ABB RAPID module: Main.mod

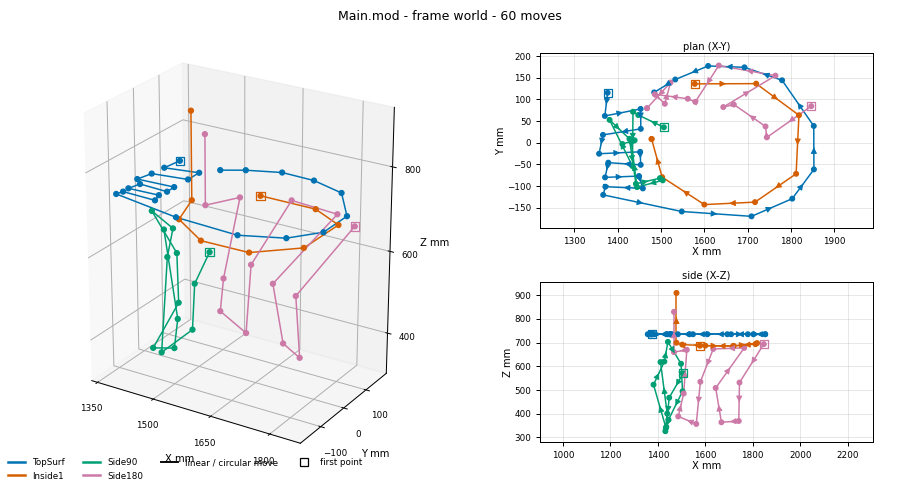
[picture p0: tool path of Main.mod in frame world, 60 of 82 moves have a stored position in this frame; points joined in program order, loops and branches not executed]
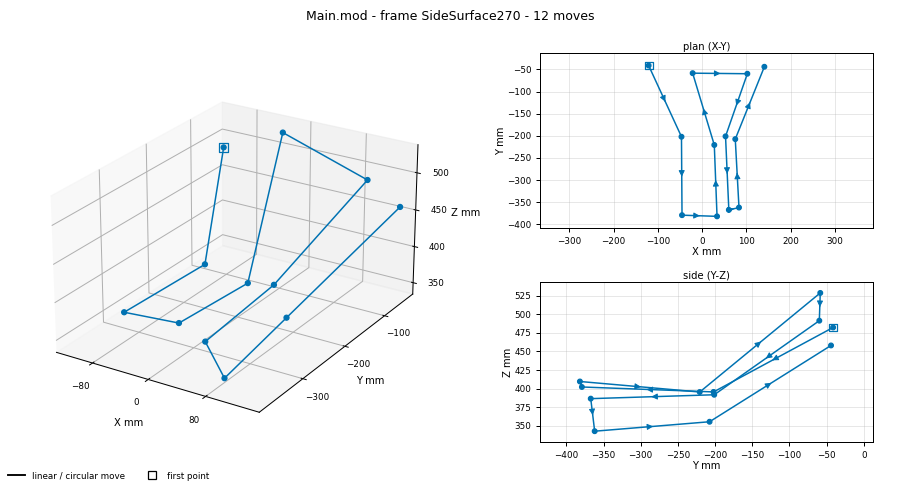
[picture p1: tool path of Main.mod in frame SideSurface270, 12 of 82 moves have a stored position in this frame; points joined in program order, loops and branches not executed]
%%%
  VERSION:1
  LANGUAGE:ENGLISH
%%%
MODULE MOD_Main

    ! -------------------------------
    ! Define customized variables here
    ! ...

	! Tool variables:
	PERS tooldata ToolRDK2 := [TRUE,[[-397.000,-4.578,191.692],[0.70710678,0.00000000,-0.70710678,0.00000001]],[1,[0,0,20],[1,0,0,0],0,0,0.005]];
	PERS tooldata ToolRDKRy15 := [TRUE,[[-327.000,-4.578,191.692],[0.60876143,0.00000000,-0.79335334,-0.00000000]],[1,[0,0,20],[1,0,0,0],0,0,0.005]];

	! Reference variables:
	PERS wobjdata SideSurface270 := [FALSE, TRUE, "", [[0,0,0],[1,0,0,0]],[[1336.130,0.000,735.410],[0.50000000,0.50000000,0.50000000,0.50000000]]];
	PERS wobjdata TopSurf2 := [FALSE, TRUE, "", [[0,0,0],[1,0,0,0]],[[1336.130,0.000,735.410],[0.50000000,0.50000000,0.50000000,0.50000000]]];
	PERS wobjdata Inside := [FALSE, TRUE, "", [[0,0,0],[1,0,0,0]],[[1336.130,0.000,735.410],[0.50000000,0.50000000,0.50000000,0.50000000]]];
	PERS wobjdata SideSurface90 := [FALSE, TRUE, "", [[0,0,0],[1,0,0,0]],[[1336.130,0.000,735.410],[0.50000000,0.50000000,0.50000000,0.50000000]]];
	PERS wobjdata SdeSurface180 := [FALSE, TRUE, "", [[0,0,0],[1,0,0,0]],[[1336.130,0.000,735.410],[0.50000000,0.50000000,0.50000000,0.50000000]]];

	PROC TopSurf()
		ConfJ \On;
		ConfL \Off;
		TT0deg;
		ToolRDK2 := [TRUE,[[-397.000,-4.578,191.692],[0.70710678,0.00000000,-0.70710678,0.00000001]],[1,[0,0,20],[1,0,0,0],0,0,0.005]];
		MoveAbsJ [[-2.762230,35.281600,-32.244600,94.063100,36.825000,84.928900],[9E+09,9E+09,9E+09,9E+09,9E+09,9E+09]],v500,z1,ToolRDK2 \WObj:=TopSurf2;
		MoveAbsJ [[3.888270,37.649400,-27.622300,84.244200,-60.438300,101.547000],[9E+09,9E+09,9E+09,9E+09,9E+09,9E+09]],v500,z1,ToolRDK2 \WObj:=TopSurf2;
		GunOn 1;
		MoveL [[115.290,-0.000,40.893],[0.66951661,0.66951663,0.22748073,-0.22748077],[-1,1,1,2],[9E+09,9E+09,9E+09,9E+09,9E+09,9E+09]],v500,z1,ToolRDK2 \WObj:=TopSurf2;
		MoveL [[61.769,-0.000,34.498],[0.66824739,0.66824741,0.23118262,-0.23118267],[0,0,1,1],[9E+09,9E+09,9E+09,9E+09,9E+09,9E+09]],v500,z1,ToolRDK2 \WObj:=TopSurf2;
		MoveL [[77.918,0.000,116.954],[0.67411479,0.67411479,0.21346957,-0.21346957],[0,0,1,1],[9E+09,9E+09,9E+09,9E+09,9E+09,9E+09]],v500,z1,ToolRDK2 \WObj:=TopSurf2;
		MoveL [[32.029,0.000,117.425],[0.67416339,0.67416339,0.21331602,-0.21331602],[0,0,1,1],[9E+09,9E+09,9E+09,9E+09,9E+09,9E+09]],v500,z1,ToolRDK2 \WObj:=TopSurf2;
		MoveL [[18.094,-0.000,30.124],[0.66795555,0.66795555,0.23202454,-0.23202454],[0,0,1,1],[9E+09,9E+09,9E+09,9E+09,9E+09,9E+09]],v500,z1,ToolRDK2 \WObj:=TopSurf2;
		MoveL [[-25.377,-0.000,21.201],[0.66687834,0.66687834,0.23510269,-0.23510270],[0,0,1,1],[9E+09,9E+09,9E+09,9E+09,9E+09,9E+09]],v500,z1,ToolRDK2 \WObj:=TopSurf2;
		MoveL [[-20.929,0.000,115.878],[0.67369753,0.67369752,0.21478279,-0.21478278],[0,0,1,1],[9E+09,9E+09,9E+09,9E+09,9E+09,9E+09]],v500,z1,ToolRDK2 \WObj:=TopSurf2;
		MoveL [[-51.029,0.000,117.232],[0.67365028,0.67365028,0.21493093,-0.21493093],[0,0,1,1],[9E+09,9E+09,9E+09,9E+09,9E+09,9E+09]],v500,z1,ToolRDK2 \WObj:=TopSurf2;
		MoveL [[-45.916,-0.000,42.441],[0.66826232,0.66826233,0.23113949,-0.23113950],[0,0,1,1],[9E+09,9E+09,9E+09,9E+09,9E+09,9E+09]],v500,z1,ToolRDK2 \WObj:=TopSurf2;
		MoveL [[-79.907,-0.000,34.972],[0.66736193,0.66736194,0.23372644,-0.23372644],[0,0,1,1],[9E+09,9E+09,9E+09,9E+09,9E+09,9E+09]],v500,z1,ToolRDK2 \WObj:=TopSurf2;
		MoveL [[-76.800,0.000,113.142],[0.67321469,0.67321469,0.21629141,-0.21629141],[0,0,1,1],[9E+09,9E+09,9E+09,9E+09,9E+09,9E+09]],v500,z1,ToolRDK2 \WObj:=TopSurf2;
		MoveL [[-105.332,0.000,122.191],[0.67370783,0.67370783,0.21475045,-0.21475045],[0,0,1,1],[9E+09,9E+09,9E+09,9E+09,9E+09,9E+09]],v500,z1,ToolRDK2 \WObj:=TopSurf2;
		MoveL [[-101.402,-0.000,35.713],[0.66719553,0.66719554,0.23420101,-0.23420104],[0,0,1,1],[9E+09,9E+09,9E+09,9E+09,9E+09,9E+09]],v500,z1,ToolRDK2 \WObj:=TopSurf2;
		MoveL [[-120.231,-0.000,30.646],[0.66659020,0.66659020,0.23591842,-0.23591844],[0,0,1,1],[9E+09,9E+09,9E+09,9E+09,9E+09,9E+09]],v500,z1,ToolRDK2 \WObj:=TopSurf2;
		MoveL [[-158.578,-0.000,211.837],[0.67989399,0.67989399,0.19427858,-0.19427858],[0,2,-1,0],[9E+09,9E+09,9E+09,9E+09,9E+09,9E+09]],v500,z1,ToolRDK2 \WObj:=TopSurf2;
		MoveL [[-169.769,-0.000,372.687],[0.68989069,0.68989069,0.15508330,-0.15508330],[0,2,-1,0],[9E+09,9E+09,9E+09,9E+09,9E+09,9E+09]],v500,z1,ToolRDK2 \WObj:=TopSurf2;
		MoveL [[-128.964,0.000,466.626],[0.69493868,0.69493868,0.13061485,-0.13061485],[0,2,-1,0],[9E+09,9E+09,9E+09,9E+09,9E+09,9E+09]],v500,z1,ToolRDK2 \WObj:=TopSurf2;
		MoveL [[-61.529,0.000,516.598],[0.69594843,0.69594843,0.12512308,-0.12512308],[0,2,-1,0],[9E+09,9E+09,9E+09,9E+09,9E+09,9E+09]],v500,z1,ToolRDK2 \WObj:=TopSurf2;
		MoveL [[38.647,0.000,516.273],[0.69521781,0.69521781,0.12912086,-0.12912086],[0,2,-1,0],[9E+09,9E+09,9E+09,9E+09,9E+09,9E+09]],v500,z1,ToolRDK2 \WObj:=TopSurf2;
		MoveL [[144.073,0.000,443.157],[0.69160511,0.69160511,0.14724934,-0.14724934],[0,0,1,1],[9E+09,9E+09,9E+09,9E+09,9E+09,9E+09]],v500,z1,ToolRDK2 \WObj:=TopSurf2;
		MoveL [[173.888,-0.000,356.448],[0.68759917,0.68759917,0.16494659,-0.16494659],[0,0,1,1],[9E+09,9E+09,9E+09,9E+09,9E+09,9E+09]],v500,z1,ToolRDK2 \WObj:=TopSurf2;
		MoveL [[177.057,0.000,272.670],[0.68344550,0.68344550,0.18138976,-0.18138976],[0,0,1,1],[9E+09,9E+09,9E+09,9E+09,9E+09,9E+09]],v500,z1,ToolRDK2 \WObj:=TopSurf2;
		MoveL [[145.838,-0.000,196.841],[0.67931130,0.67931130,0.19630627,-0.19630627],[0,0,1,1],[9E+09,9E+09,9E+09,9E+09,9E+09,9E+09]],v500,z1,ToolRDK2 \WObj:=TopSurf2;
		GunOn 0;
		MoveL [[116.077,0.000,148.259],[0.67637750,0.67637750,0.20618797,-0.20618797],[0,0,1,1],[9E+09,9E+09,9E+09,9E+09,9E+09,9E+09]],v500,z1,ToolRDK2 \WObj:=TopSurf2;
	ENDPROC

	PROC TT0deg()
		ConfJ \On;
		ConfL \Off;
		MoveAbsJ [[0.000000,0.000000,0.000000,0.000000,0.000000,0.000000],[9E+09,9E+09,9E+09,9E+09,9E+09,9E+09]],v500,z1,ToolRDK2 \WObj:=TopSurf2;
	ENDPROC

	PROC Inside1()
		ConfJ \On;
		ConfL \Off;
		TT0deg;
		MoveAbsJ [[-5.345720,35.456100,-20.669400,-15.550700,88.287700,-47.645500],[9E+09,9E+09,9E+09,9E+09,9E+09,9E+09]],v500,z1,ToolRDKRy15 \WObj:=Inside;
		GunOn 1;
		MoveL [[135.749,-48.253,241.842],[0.26164486,-0.62731638,0.51686708,-0.52044649],[-1,-1,-2,0],[9E+09,9E+09,9E+09,9E+09,9E+09,9E+09]],v100,z1,ToolRDKRy15 \WObj:=Inside;
		MoveL [[136.293,-48.875,383.457],[0.53837192,-0.31876420,0.47937269,-0.61542415],[-1,-1,3,0],[9E+09,9E+09,9E+09,9E+09,9E+09,9E+09]],v100,z1,ToolRDKRy15 \WObj:=Inside;
		MoveL [[63.451,-37.348,482.087],[0.60930435,-0.14318770,0.26615634,-0.73308001],[0,-1,3,0],[9E+09,9E+09,9E+09,9E+09,9E+09,9E+09]],v100,z1,ToolRDKRy15 \WObj:=Inside;
		MoveL [[-71.616,-41.647,475.560],[0.73598605,0.22123419,-0.09604572,-0.63257820],[-1,0,0,0],[9E+09,9E+09,9E+09,9E+09,9E+09,9E+09]],v100,z1,ToolRDKRy15 \WObj:=Inside;
		MoveL [[-136.962,-50.085,380.769],[0.64868094,0.45794626,-0.34884692,-0.49779925],[-1,0,0,0],[9E+09,9E+09,9E+09,9E+09,9E+09,9E+09]],v100,z1,ToolRDKRy15 \WObj:=Inside;
		MoveL [[-142.620,-47.996,263.919],[0.46214789,0.64281008,-0.47460814,-0.38465783],[-1,0,1,0],[9E+09,9E+09,9E+09,9E+09,9E+09,9E+09]],v100,z1,ToolRDKRy15 \WObj:=Inside;
		MoveL [[-79.374,-43.840,166.588],[0.24696012,0.71987130,-0.64178535,-0.09437996],[-1,0,1,0],[9E+09,9E+09,9E+09,9E+09,9E+09,9E+09]],v100,z1,ToolRDKRy15 \WObj:=Inside;
		MoveL [[8.609,-35.875,142.282],[0.04464887,0.71177006,-0.69465400,0.09405146],[-1,0,2,0],[9E+09,9E+09,9E+09,9E+09,9E+09,9E+09]],v100,z1,ToolRDKRy15 \WObj:=Inside;
		GunOn 0;
		MoveL [[8.609,174.125,142.282],[0.04464720,0.71176897,-0.69465549,0.09404953],[0,3,4,0],[9E+09,9E+09,9E+09,9E+09,9E+09,9E+09]],v100,z1,ToolRDKRy15 \WObj:=Inside;
	ENDPROC

	PROC Side90()
		ConfJ \On;
		ConfL \Off;
		TT90deg;
		ToolRDK2 := [TRUE,[[-397.000,-4.578,191.692],[0.70710678,0.00000000,-0.70710678,0.00000001]],[1,[0,0,20],[1,0,0,0],0,0,0.005]];
		MoveAbsJ [[2.579840,12.805000,8.075260,-0.378023,73.507000,3.846430],[9E+09,9E+09,9E+09,9E+09,9E+09,9E+09]],v100,z1,ToolRDK2 \WObj:=SideSurface90;
		MoveL [[35.648,-164.659,170.589],[0.70282661,0.03396154,0.01983662,-0.71027310],[0,-1,0,0],[9E+09,9E+09,9E+09,9E+09,9E+09,9E+09]],v100,z1,ToolRDK2 \WObj:=SideSurface90;
		GunOn 1;
		MoveL [[63.939,-267.719,111.565],[0.70282661,0.03396154,0.01983662,-0.71027310],[0,-1,0,0],[9E+09,9E+09,9E+09,9E+09,9E+09,9E+09]],v100,z1,ToolRDK2 \WObj:=SideSurface90;
		MoveL [[71.496,-390.187,99.400],[0.70282661,0.03396154,0.01983662,-0.71027310],[0,-1,0,0],[9E+09,9E+09,9E+09,9E+09,9E+09,9E+09]],v100,z1,ToolRDK2 \WObj:=SideSurface90;
		MoveL [[-53.749,-395.227,98.058],[0.70282661,0.03396154,0.01983662,-0.71027310],[-1,-1,0,0],[9E+09,9E+09,9E+09,9E+09,9E+09,9E+09]],v100,z1,ToolRDK2 \WObj:=SideSurface90;
		MoveL [[52.643,-212.764,45.439],[0.70282661,0.03396154,0.01983662,-0.71027310],[0,-1,0,0],[9E+09,9E+09,9E+09,9E+09,9E+09,9E+09]],v100,z1,ToolRDK2 \WObj:=SideSurface90;
		MoveL [[8.984,-115.328,91.184],[0.70282661,0.03396154,0.01983662,-0.71027310],[0,-1,0,0],[9E+09,9E+09,9E+09,9E+09,9E+09,9E+09]],v100,z1,ToolRDK2 \WObj:=SideSurface90;
		MoveL [[-94.720,-32.255,106.179],[0.70282661,0.03396154,0.01983662,-0.71027310],[-1,-1,-1,0],[9E+09,9E+09,9E+09,9E+09,9E+09,9E+09]],v100,z1,ToolRDK2 \WObj:=SideSurface90;
		MoveL [[-81.740,-124.404,161.457],[0.70282661,0.03396154,0.01983662,-0.71027310],[-1,-1,-1,0],[9E+09,9E+09,9E+09,9E+09,9E+09,9E+09]],v100,z1,ToolRDK2 \WObj:=SideSurface90;
		MoveL [[-86.756,-240.544,167.927],[0.70282661,0.03396154,0.01983662,-0.71027310],[-1,-1,-1,0],[9E+09,9E+09,9E+09,9E+09,9E+09,9E+09]],v100,z1,ToolRDK2 \WObj:=SideSurface90;
		MoveL [[-102.328,-360.623,108.637],[0.70282661,0.03396154,0.01983662,-0.71027310],[-1,-1,-1,0],[9E+09,9E+09,9E+09,9E+09,9E+09,9E+09]],v100,z1,ToolRDK2 \WObj:=SideSurface90;
		MoveL [[1.978,-408.957,95.385],[0.70282661,0.03396154,0.01983662,-0.71027310],[0,-1,0,0],[9E+09,9E+09,9E+09,9E+09,9E+09,9E+09]],v100,z1,ToolRDK2 \WObj:=SideSurface90;
		MoveL [[5.518,-334.746,103.233],[0.70282661,0.03396154,0.01983662,-0.71027310],[0,-1,0,0],[9E+09,9E+09,9E+09,9E+09,9E+09,9E+09]],v100,z1,ToolRDK2 \WObj:=SideSurface90;
		MoveL [[-2.937,-117.398,74.861],[0.70282661,0.03396154,0.01983662,-0.71027310],[0,-1,0,0],[9E+09,9E+09,9E+09,9E+09,9E+09,9E+09]],v100,z1,ToolRDK2 \WObj:=SideSurface90;
		GunOn 0;
	ENDPROC

	PROC TT90deg()
		ConfJ \On;
		ConfL \Off;
		MoveAbsJ [[90.000000,0.000000,0.000000,0.000000,0.000000,0.000000],[9E+09,9E+09,9E+09,9E+09,9E+09,9E+09]],v100,z1,ToolRDK2 \WObj:=SideSurface90;
	ENDPROC

	PROC Side180()
		ConfJ \On;
		ConfL \Off;
		TT180deg;
		ToolRDK2 := [TRUE,[[-397.000,-4.578,191.692],[0.70710678,0.00000000,-0.70710678,0.00000001]],[1,[0,0,20],[1,0,0,0],0,0,0.005]];
		MoveAbsJ [[22.186600,36.517800,-32.653500,15.382700,96.981900,81.677400],[9E+09,9E+09,9E+09,9E+09,9E+09,9E+09]],v100,z1,ToolRDK2 \WObj:=SdeSurface180;
		MoveL [[84.401,-41.748,510.527],[0.27194744,0.74951284,-0.59519100,-0.10011380],[-1,-1,-1,0],[9E+09,9E+09,9E+09,9E+09,9E+09,9E+09]],v100,z1,ToolRDK2 \WObj:=SdeSurface180;
		GunOn 1;
		MoveL [[12.341,-203.862,408.074],[0.19866001,0.68168548,-0.69934461,-0.08219625],[-1,-1,-1,0],[9E+09,9E+09,9E+09,9E+09,9E+09,9E+09]],v100,z1,ToolRDK2 \WObj:=SdeSurface180;
		MoveL [[37.555,-365.927,404.980],[0.30278680,0.66474465,-0.62196033,-0.28213480],[-1,-1,-1,0],[9E+09,9E+09,9E+09,9E+09,9E+09,9E+09]],v100,z1,ToolRDK2 \WObj:=SdeSurface180;
		MoveL [[88.260,-371.346,331.859],[0.56338823,0.56604743,-0.42378097,-0.42730985],[0,0,-3,0],[9E+09,9E+09,9E+09,9E+09,9E+09,9E+09]],v100,z1,ToolRDK2 \WObj:=SdeSurface180;
		MoveL [[82.260,-226.787,307.601],[0.57594149,0.55309259,-0.44055486,-0.41023334],[0,0,-3,0],[9E+09,9E+09,9E+09,9E+09,9E+09,9E+09]],v100,z1,ToolRDK2 \WObj:=SdeSurface180;
		MoveL [[154.718,-57.664,427.892],[0.40312792,0.63471100,-0.54999996,-0.36349672],[-1,-1,-1,0],[9E+09,9E+09,9E+09,9E+09,9E+09,9E+09]],v100,z1,ToolRDK2 \WObj:=SdeSurface180;
		MoveL [[178.045,-62.096,297.332],[0.56841264,0.56098553,-0.43045933,-0.42060323],[0,0,-3,0],[9E+09,9E+09,9E+09,9E+09,9E+09,9E+09]],v100,z1,ToolRDK2 \WObj:=SdeSurface180;
		MoveL [[94.348,-200.545,243.065],[0.54952518,0.57922797,-0.40557979,-0.44499672],[0,0,-3,0],[9E+09,9E+09,9E+09,9E+09,9E+09,9E+09]],v100,z1,ToolRDK2 \WObj:=SdeSurface180;
		MoveL [[101.429,-378.373,225.720],[0.52959167,0.59636781,-0.37992820,-0.46854313],[0,0,-3,0],[9E+09,9E+09,9E+09,9E+09,9E+09,9E+09]],v100,z1,ToolRDK2 \WObj:=SdeSurface180;
		MoveL [[111.805,-346.628,149.664],[0.54531210,0.58302000,-0.40010958,-0.45014965],[0,0,-3,0],[9E+09,9E+09,9E+09,9E+09,9E+09,9E+09]],v100,z1,ToolRDK2 \WObj:=SdeSurface180;
		MoveL [[89.794,-249.802,172.785],[0.55734821,0.57192725,-0.41581153,-0.43515856],[0,0,-3,0],[9E+09,9E+09,9E+09,9E+09,9E+09,9E+09]],v100,z1,ToolRDK2 \WObj:=SdeSurface180;
		MoveL [[138.848,-65.706,185.941],[0.49595548,0.52244183,-0.46707769,-0.51275835],[0,0,-3,0],[9E+09,9E+09,9E+09,9E+09,9E+09,9E+09]],v100,z1,ToolRDK2 \WObj:=SdeSurface180;
		MoveL [[79.680,-75.532,131.744],[0.70566624,0.20024459,-0.17913763,-0.65562716],[0,0,-4,0],[9E+09,9E+09,9E+09,9E+09,9E+09,9E+09]],v100,z1,ToolRDK2 \WObj:=SdeSurface180;
		MoveL [[79.680,94.467,131.744],[0.70566463,0.20024809,-0.17913633,-0.65562818],[0,0,0,0],[9E+09,9E+09,9E+09,9E+09,9E+09,9E+09]],v100,z1,ToolRDK2 \WObj:=SdeSurface180;
		GunOn 0;
	ENDPROC

	PROC TT180deg()
		ConfJ \On;
		ConfL \Off;
		MoveAbsJ [[180.000000,0.000000,0.000000,0.000000,0.000000,0.000000],[9E+09,9E+09,9E+09,9E+09,9E+09,9E+09]],v100,z1,ToolRDK2 \WObj:=SdeSurface180;
	ENDPROC

	PROC Side270()
		ConfJ \On;
		ConfL \Off;
		TT270deg;
		SideSurface270 := [FALSE, TRUE, "", [[0,0,0],[1,0,0,0]],[[1336.130,0.000,735.410],[0.50000000,0.50000000,0.50000000,0.50000000]]];
		ToolRDK2 := [TRUE,[[-397.000,-4.578,191.692],[0.70710678,0.00000000,-0.70710678,0.00000001]],[1,[0,0,20],[1,0,0,0],0,0,0.005]];
		MoveAbsJ [[17.239800,6.188030,12.545200,5.893900,70.141500,47.412000],[9E+09,9E+09,9E+09,9E+09,9E+09,9E+09]],v100,z1,ToolRDK2 \WObj:=SideSurface270;
		MoveL [[-120.767,-41.372,482.237],[0.21739829,-0.63519472,0.69915740,-0.24585480],[0,-2,-2,1],[9E+09,9E+09,9E+09,9E+09,9E+09,9E+09]],v100,z1,ToolRDK2 \WObj:=SideSurface270;
		GunOn 1;
		MoveL [[-46.657,-202.048,395.599],[0.18859986,-0.66328159,0.67980013,-0.24971865],[0,0,0,0],[9E+09,9E+09,9E+09,9E+09,9E+09,9E+09]],v100,z1,ToolRDK2 \WObj:=SideSurface270;
		MoveL [[-45.433,-379.054,402.243],[0.10607148,-0.70258822,0.68574611,-0.15770515],[0,0,0,0],[9E+09,9E+09,9E+09,9E+09,9E+09,9E+09]],v100,z1,ToolRDK2 \WObj:=SideSurface270;
		MoveL [[33.587,-381.726,409.620],[0.01983662,0.71027310,-0.70282661,0.03396154],[-1,-1,0,0],[9E+09,9E+09,9E+09,9E+09,9E+09,9E+09]],v100,z1,ToolRDK2 \WObj:=SideSurface270;
		MoveL [[27.391,-220.636,395.484],[0.01983662,0.71027310,-0.70282661,0.03396154],[-1,-1,0,0],[9E+09,9E+09,9E+09,9E+09,9E+09,9E+09]],v100,z1,ToolRDK2 \WObj:=SideSurface270;
		MoveL [[-21.445,-58.617,528.661],[0.04513872,-0.70911484,0.69678436,-0.09803156],[0,-1,0,0],[9E+09,9E+09,9E+09,9E+09,9E+09,9E+09]],v100,z1,ToolRDK2 \WObj:=SideSurface270;
		MoveL [[101.993,-59.897,491.361],[0.26329516,0.65992995,-0.67147736,-0.21044306],[-1,-1,-1,0],[9E+09,9E+09,9E+09,9E+09,9E+09,9E+09]],v100,z1,ToolRDK2 \WObj:=SideSurface270;
		MoveL [[52.755,-201.170,391.792],[0.26329516,0.65992995,-0.67147736,-0.21044306],[-1,-1,-1,0],[9E+09,9E+09,9E+09,9E+09,9E+09,9E+09]],v100,z1,ToolRDK2 \WObj:=SideSurface270;
		MoveL [[60.207,-367.169,386.569],[0.26329516,0.65992995,-0.67147736,-0.21044306],[-1,-1,-1,0],[9E+09,9E+09,9E+09,9E+09,9E+09,9E+09]],v100,z1,ToolRDK2 \WObj:=SideSurface270;
		MoveL [[83.108,-361.868,342.805],[0.26329516,0.65992995,-0.67147736,-0.21044306],[-1,-1,-1,0],[9E+09,9E+09,9E+09,9E+09,9E+09,9E+09]],v100,z1,ToolRDK2 \WObj:=SideSurface270;
		MoveL [[74.721,-207.428,355.509],[0.26329516,0.65992995,-0.67147736,-0.21044306],[-1,-1,-1,0],[9E+09,9E+09,9E+09,9E+09,9E+09,9E+09]],v100,z1,ToolRDK2 \WObj:=SideSurface270;
		MoveL [[140.381,-44.162,458.070],[0.26329516,0.65992995,-0.67147736,-0.21044306],[-1,-1,-1,0],[9E+09,9E+09,9E+09,9E+09,9E+09,9E+09]],v100,z1,ToolRDK2 \WObj:=SideSurface270;
		GunOn 0;
	ENDPROC

	PROC TT270deg()
		ConfJ \On;
		ConfL \Off;
		MoveAbsJ [[270.000000,0.000000,0.000000,0.000000,0.000000,0.000000],[9E+09,9E+09,9E+09,9E+09,9E+09,9E+09]],v100,z1,ToolRDK2 \WObj:=SideSurface270;
	ENDPROC

	PROC Main()
		ConfJ \On;
		ConfL \Off;
		! Program generated by VerticalBot Studio for ABB IRB 2600-12/1.85 on 25/10/2026 12:00:00
		! Using nominal kinematics.
		TopSurf;
		Inside1;
		Side0;
		Side90;
		Side180;
		Side270;
	ENDPROC

ENDMODULE
